TYPE (* logiBUS 2 CAN DI Struct Octal *)
  (* Version 1.0, 2026-05-28, franz *)
  PACKAGE logiBUS::io::DI_CAN;
  IMPORT logiBUS::io::DI_CAN::logiBUS_2_CAN_DI_S;
  logiBUS_2_CAN_DI_S_Octal : STRUCT
    Port1 : logiBUS_2_CAN_DI_S := (Pin := 255);
    Port2 : logiBUS_2_CAN_DI_S := (Pin := 255);
    Port3 : logiBUS_2_CAN_DI_S := (Pin := 255);
    Port4 : logiBUS_2_CAN_DI_S := (Pin := 255);
    Port5 : logiBUS_2_CAN_DI_S := (Pin := 255);
    Port6 : logiBUS_2_CAN_DI_S := (Pin := 255);
    Port7 : logiBUS_2_CAN_DI_S := (Pin := 255);
    Port8 : logiBUS_2_CAN_DI_S := (Pin := 255);
  END_STRUCT;
END_TYPE
